(*
SPDX-FileCopyrightText: © 2026 Oleksandr Tiutyk <trofimich@gmail.com>
SPDX-License-Identifier: MIT
License: https://opensource.org/license/mit
*)

(*!
<summary>Provides finite bounds for UnsignedInt64 values.</summary>
<description>
MIN_VALUE and MAX_VALUE describe the represented integer range; constants perform no conversion or runtime
validation. Additional named bounds, where declared, describe narrower representations.
</description>
*)

{attribute 'no_explicit_call' := 'do not call this function block directly'}
PROGRAM UnsignedInt64
VAR CONSTANT
	ZERO : ULINT := 0;
	MIN_VALUE : ULINT := 0;
	MAX_VALUE : ULINT := ULINT#16#FFFFFFFFFFFFFFFF;
END_VAR
VAR
	{attribute 'hide'} 
	_ClassName : STRING := __POUNAME();
END_VAR

{attribute 'monitoring' := 'call'}
PROPERTY ClassName : REFERENCE TO STRING
GET
ClassName REF= _ClassName;
END_GET
END_PROPERTY

(*!
<summary>Provides the library namespace used in diagnostics.</summary>
<description>
Borrowed read-only reference to the compiler-initialized library namespace; no ownership transfer.
</description>
*)
{attribute 'monitoring' := 'call'}
PROPERTY NamespaceName : REFERENCE TO STRING
GET
NamespaceName REF= CurrentNamespace.Name;
END_GET
END_PROPERTY

END_PROGRAM

(* stored: Version 1.1.0.1
   POU UnsignedInt64: Id {58df88cf-50aa-4336-8cc5-101184ba5ae9}, SpecialFunc None
   Property ClassName: Id {c9902b8b-4441-4db4-9836-61de8230deed}
   Get Get: Id {72636f1c-39cf-4e74-8ad7-9656e317c009}
   Property NamespaceName: Id {83f4fb94-795a-4980-a2a3-17badd4fcbbb}
   Get Get: Id {b608a452-9359-4c01-bfd0-24267a1c3c3b} *)
